DATA_BLOCK "FRK_Decisions"
{ S7_Optimized_Access := 'TRUE' }
VERSION : 0.1
NON_RETAIN
VAR
    Slots {ExternalAccessible := 'False'; ExternalVisible := 'False'; ExternalWritable := 'False'} : Array[1..2] of "FRK_DecisionSlot";
    EmptyRequest {ExternalAccessible := 'False'; ExternalVisible := 'False'; ExternalWritable := 'False'} : "ST_DecisionRequest";
END_VAR
BEGIN
END_DATA_BLOCK
